(* IEC 61131-3 sources: llm-plc-st-eval/data/processed_definitivo/qwen2.5-coder_14b/A2/zero_shot, 3 files *)

(* ---- ejec_1.st ---- *)
FUNCTION_BLOCK FB_Batch
VAR_INPUT
    nivelA, nivelB, nivelVacio, btnInicio, btnAbort : BOOL;
    temp : REAL;
END_VAR

VAR_OUTPUT
    vA, vB, calentador, mezclador, vDescarga : BOOL;
    fase : INT;
END_VAR

VAR
    timerMezclador : TON;
    estado : INT := 0; // 0: reposo, 1: fase 1, 2: fase 2, 3: fase 3, 4: fase 4, 5: fase 5
END_VAR

METHOD StartBatch : VOID
    IF btnInicio AND estado = 0 THEN
        estado := 1;
    END_IF;
END_METHOD

METHOD AbortBatch : VOID
    IF btnAbort THEN
        vA := FALSE;
        vB := FALSE;
        calentador := FALSE;
        mezclador := FALSE;

        IF nivelVacio THEN
            estado := 0;
        ELSE
            estado := 5;
        END_IF;
    END_IF;
END_METHOD

METHOD UpdateBatch : VOID
    CASE estado OF
        0: // Reposo
            fase := 0;
            vA := FALSE;
            vB := FALSE;
            calentador := FALSE;
            mezclador := FALSE;
            vDescarga := FALSE;

        1: // Fase 1: Dosificar componente A
            fase := 1;
            vA := TRUE;
            IF nivelA THEN
                vA := FALSE;
                estado := 2;
            END_IF;

        2: // Fase 2: Dosificar componente B
            fase := 2;
            vB := TRUE;
            IF nivelB THEN
                vB := FALSE;
                estado := 3;
            END_IF;

        3: // Fase 3: Calentar
            fase := 3;
            calentador := TRUE;
            IF temp >= 60.0 THEN
                calentador := FALSE;
                estado := 4;
            END_IF;

        4: // Fase 4: Mezclar
            fase := 4;
            mezclador := TRUE;
            timerMezclador(IN := TRUE, PT := T#120S);
            IF timerMezclador.Q THEN
                mezclador := FALSE;
                timerMezclador(IN := FALSE);
                estado := 5;
            END_IF;

        5: // Fase 5: Descargar
            fase := 5;
            vDescarga := TRUE;
            IF nivelVacio THEN
                vDescarga := FALSE;
                estado := 0;
            END_IF;
    END_CASE;
END_METHOD

METHOD Execute : VOID
    StartBatch();
    AbortBatch();
    UpdateBatch();
END_METHOD

(* ---- ejec_2.st ---- *)
FUNCTION_BLOCK FB_Batch
VAR_INPUT
    nivelA, nivelB, nivelVacio, btnInicio, btnAbort : BOOL;
    temp : REAL;
END_VAR

VAR_OUTPUT
    vA, vB, calentador, mezclador, vDescarga : BOOL;
    fase : INT;
END_VAR

VAR
    timerMezclador : TON;
    estado : INT := 0; // 0: reposo, 1: dosificar A, 2: dosificar B, 3: calentar, 4: mezclar, 5: descargar
    timerMezcladorActive : BOOL := FALSE;
END_VAR

METHOD StartBatch : BOOL
    IF btnInicio AND estado = 0 THEN
        estado := 1;
        RETURN TRUE;
    END_IF
    RETURN FALSE;
END_METHOD

METHOD AbortBatch : BOOL
    IF btnAbort AND estado > 0 THEN
        vA := FALSE;
        vB := FALSE;
        calentador := FALSE;
        mezclador := FALSE;
        IF NOT nivelVacio THEN
            estado := 5;
        ELSE
            estado := 0;
        END_IF
        RETURN TRUE;
    END_IF
    RETURN FALSE;
END_METHOD

METHOD UpdateBatch : BOOL
    CASE estado OF
        0: // Reposo
            vA := FALSE;
            vB := FALSE;
            calentador := FALSE;
            mezclador := FALSE;
            vDescarga := FALSE;
            fase := 0;
        1: // Dosificar A
            vA := TRUE;
            vB := FALSE;
            calentador := FALSE;
            mezclador := FALSE;
            vDescarga := FALSE;
            fase := 1;
            IF nivelA THEN
                vA := FALSE;
                estado := 2;
            END_IF;
        2: // Dosificar B
            vA := FALSE;
            vB := TRUE;
            calentador := FALSE;
            mezclador := FALSE;
            vDescarga := FALSE;
            fase := 2;
            IF nivelB THEN
                vB := FALSE;
                estado := 3;
            END_IF;
        3: // Calentar
            vA := FALSE;
            vB := FALSE;
            calentador := TRUE;
            mezclador := FALSE;
            vDescarga := FALSE;
            fase := 3;
            IF temp >= 60.0 THEN
                calentador := FALSE;
                estado := 4;
            END_IF;
        4: // Mezclar
            vA := FALSE;
            vB := FALSE;
            calentador := FALSE;
            mezclador := TRUE;
            vDescarga := FALSE;
            fase := 4;
            IF NOT timerMezcladorActive THEN
                timerMezclador(IN := TRUE, PT := T#120S);
                timerMezcladorActive := TRUE;
            END_IF;
            IF timerMezclador.Q THEN
                mezclador := FALSE;
                timerMezcladorActive := FALSE;
                estado := 5;
            END_IF;
        5: // Descargar
            vA := FALSE;
            vB := FALSE;
            calentador := FALSE;
            mezclador := FALSE;
            vDescarga := TRUE;
            fase := 5;
            IF nivelVacio THEN
                vDescarga := FALSE;
                estado := 0;
            END_IF;
    END_CASE
    RETURN TRUE;
END_METHOD

METHOD Execute : BOOL
    IF AbortBatch() THEN
        RETURN TRUE;
    END_IF;
    IF StartBatch() THEN
        RETURN TRUE;
    END_IF;
    IF UpdateBatch() THEN
        RETURN TRUE;
    END_IF;
    RETURN FALSE;
END_METHOD

METHOD Reset : BOOL
    estado := 0;
    RETURN TRUE;
END_METHOD
END_FUNCTION_BLOCK

(* ---- ejec_3.st ---- *)
FUNCTION_BLOCK FB_Batch
VAR_INPUT
    nivelA, nivelB, nivelVacio, btnInicio, btnAbort : BOOL;
    temp : REAL;
END_VAR

VAR_OUTPUT
    vA, vB, calentador, mezclador, vDescarga : BOOL;
    fase : INT;
END_VAR

VAR
    timerMezclador : TON;
    estado : INT := 0; // 0: reposo, 1: dosificar A, 2: dosificar B, 3: calentar, 4: mezclar, 5: descargar
END_VAR

METHOD StartBatch : BOOL
VAR
    started : BOOL := FALSE;
END_VAR
    IF btnInicio AND estado = 0 THEN
        estado := 1;
        started := TRUE;
    END_IF
    StartBatch := started;
END_METHOD

METHOD AbortBatch : BOOL
VAR
    aborted : BOOL := FALSE;
END_VAR
    IF btnAbort AND estado > 0 THEN
        vA := FALSE;
        vB := FALSE;
        calentador := FALSE;
        mezclador := FALSE;
        IF NOT nivelVacio THEN
            estado := 5;
        ELSE
            estado := 0;
        END_IF
        aborted := TRUE;
    END_IF
    AbortBatch := aborted;
END_METHOD

METHOD UpdateBatch : BOOL
VAR
    updated : BOOL := FALSE;
END_VAR
    CASE estado OF
        0: // reposo
            vA := FALSE;
            vB := FALSE;
            calentador := FALSE;
            mezclador := FALSE;
            vDescarga := FALSE;
            fase := 0;
        1: // dosificar A
            vA := TRUE;
            vB := FALSE;
            calentador := FALSE;
            mezclador := FALSE;
            vDescarga := FALSE;
            fase := 1;
            IF nivelA THEN
                vA := FALSE;
                estado := 2;
            END_IF;
        2: // dosificar B
            vA := FALSE;
            vB := TRUE;
            calentador := FALSE;
            mezclador := FALSE;
            vDescarga := FALSE;
            fase := 2;
            IF nivelB THEN
                vB := FALSE;
                estado := 3;
            END_IF;
        3: // calentar
            vA := FALSE;
            vB := FALSE;
            calentador := TRUE;
            mezclador := FALSE;
            vDescarga := FALSE;
            fase := 3;
            IF temp >= 60.0 THEN
                calentador := FALSE;
                estado := 4;
            END_IF;
        4: // mezclar
            vA := FALSE;
            vB := FALSE;
            calentador := FALSE;
            mezclador := TRUE;
            vDescarga := FALSE;
            fase := 4;
            timerMezclador(IN := TRUE, PT := T#120S);
            IF timerMezclador.Q THEN
                mezclador := FALSE;
                estado := 5;
            END_IF;
        5: // descargar
            vA := FALSE;
            vB := FALSE;
            calentador := FALSE;
            mezclador := FALSE;
            vDescarga := TRUE;
            fase := 5;
            IF nivelVacio THEN
                vDescarga := FALSE;
                estado := 0;
            END_IF;
    END_CASE
    updated := TRUE;
    UpdateBatch := updated;
END_METHOD

METHOD Execute : BOOL
VAR
    executed : BOOL := FALSE;
END_VAR
    IF StartBatch() OR AbortBatch() OR UpdateBatch() THEN
        executed := TRUE;
    END_IF
    Execute := executed;
END_METHOD

// Main execution
Execute();
